FUNCTION_BLOCK basicPreparadorVibropac (* Preparador de polimero Vibropac VIB-3000 - logica (Modbus TCP Inovaisa) *)
  (* Standard: 61499-2 *)
  (* Version 1.0, 19/10/2026, Hidryco, Hidryco, 1.0: liga/desliga ciclo remoto (4001, reenvio a cada 5 s), reset 4002 por 3 s, leitura 4005..4019, modo automatico/manual, cfgHabilitada *)
  PACKAGE Hidryco.HidrycoLib;
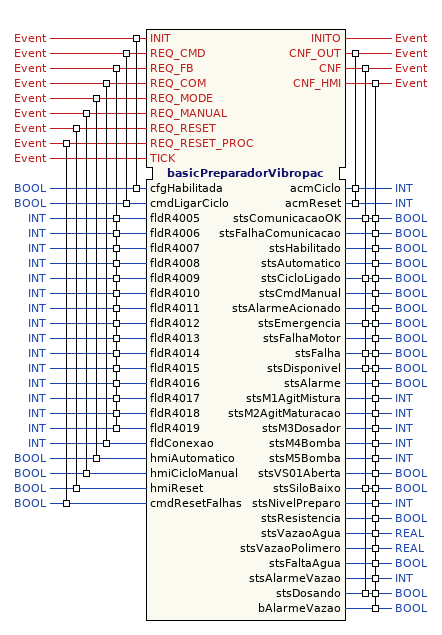
  EVENT_INPUT
    INIT WITH cfgHabilitada; (* Inicializacao (configuracao da instancia) *)
    REQ_CMD WITH cmdLigarCiclo; (* Processo: liga/desliga o ciclo (automatico) *)
    REQ_FB WITH fldR4005, fldR4006, fldR4007, fldR4008, fldR4009, fldR4010, fldR4011, fldR4012, fldR4013, fldR4014, fldR4015, fldR4016, fldR4017, fldR4018, fldR4019; (* Leitura Modbus 4005..4019 *)
    REQ_COM WITH fldConexao; (* Status da conexao Modbus (connStatusInt) *)
    REQ_MODE WITH hmiAutomatico; (* IHM: modo *)
    REQ_MANUAL WITH hmiCicloManual; (* IHM: liga/desliga o ciclo em manual *)
    REQ_RESET WITH hmiReset; (* IHM: reset *)
    REQ_RESET_PROC WITH cmdResetFalhas; (* Processo: reset *)
    TICK; (* Base de tempo de 1 s *)
  END_EVENT
  EVENT_OUTPUT
    INITO; (* Inicializacao concluida *)
    CNF_OUT WITH acmCiclo, acmReset; (* Escrita Modbus 4001 (ciclo) e 4002 (reset) *)
    CNF WITH stsComunicacaoOK, stsDisponivel, stsCicloLigado, stsFalha, stsEmergencia, stsDosando, stsSiloBaixo; (* Status para o processo (na mudanca e a cada 1 s) *)
    CNF_HMI WITH stsComunicacaoOK, stsFalhaComunicacao, stsHabilitado, stsAutomatico, stsCicloLigado, stsCmdManual, stsAlarmeAcionado, stsEmergencia, stsFalhaMotor, stsFalha, stsDisponivel, stsAlarme, stsM1AgitMistura, stsM2AgitMaturacao, stsM3Dosador, stsM4Bomba, stsM5Bomba, stsVS01Aberta, stsSiloBaixo, stsNivelPreparo, stsResistencia, stsVazaoAgua, stsVazaoPolimero, stsFaltaAgua, stsAlarmeVazao, stsDosando, bAlarmeVazao; (* Status para a IHM e alarmes *)
  END_EVENT
  VAR_INPUT
    cfgHabilitada : BOOL := TRUE; (* FALSE = instancia desabilitada (equipamento futuro): sem alarme e nunca disponivel *)
    cmdLigarCiclo : BOOL; (* Processo: TRUE = ciclo remoto ligado *)
    fldR4005 : INT; (* Registro 4005: alarme acionado (0/1) *)
    fldR4006 : INT; (* Registro 4006: emergencia (0/1) *)
    fldR4007 : INT; (* Registro 4007: status M1 agitador do tanque de mistura (0 parado, 1 funcionando, 2 falha) *)
    fldR4008 : INT; (* Registro 4008: status M2 agitador do tanque de maturacao (0 parado, 1 funcionando, 2 falha) *)
    fldR4009 : INT; (* Registro 4009: status M3 dosador volumetrico (0 parado, 1 funcionando, 2 falha) *)
    fldR4010 : INT; (* Registro 4010: status M4 bomba dosadora M4 (0 parado, 1 funcionando, 2 falha) *)
    fldR4011 : INT; (* Registro 4011: status M5 bomba dosadora M5 (0 parado, 1 funcionando, 2 falha) *)
    fldR4012 : INT; (* Registro 4012: ver tabela Modbus *)
    fldR4013 : INT; (* Registro 4013: ver tabela Modbus *)
    fldR4014 : INT; (* Registro 4014: ver tabela Modbus *)
    fldR4015 : INT; (* Registro 4015: ver tabela Modbus *)
    fldR4016 : INT; (* Registro 4016: ver tabela Modbus *)
    fldR4017 : INT; (* Registro 4017: ver tabela Modbus *)
    fldR4018 : INT; (* Registro 4018: ver tabela Modbus *)
    fldR4019 : INT; (* Registro 4019: ver tabela Modbus *)
    fldConexao : INT; (* connStatusInt (1 = online) *)
    hmiAutomatico : BOOL; (* IHM: TRUE = automatico *)
    hmiCicloManual : BOOL; (* IHM: TRUE = liga o ciclo (manual) *)
    hmiReset : BOOL; (* IHM: reset *)
    cmdResetFalhas : BOOL; (* Processo: reset (vale com TRUE) *)
  END_VAR
  VAR_OUTPUT
    acmCiclo : INT; (* Registro 4001: 1 liga ciclo remoto, 0 desliga *)
    acmReset : INT; (* Registro 4002: 1 reseta falhas (pulso de 3 s) *)
    stsComunicacaoOK : BOOL; (* Comunicacao Modbus com o CLP do skid OK *)
    stsFalhaComunicacao : BOOL; (* Falha de comunicacao com o CLP do skid *)
    stsHabilitado : BOOL; (* Instancia habilitada (FALSE = equipamento futuro) *)
    stsAutomatico : BOOL; (* Ciclo comandado pelo processo (automatico) *)
    stsCicloLigado : BOOL; (* Comando de ciclo remoto ligado (4001 = 1) *)
    stsCmdManual : BOOL; (* Comando manual de ciclo (modo manual) *)
    stsAlarmeAcionado : BOOL; (* Alarme acionado no skid (4005) *)
    stsEmergencia : BOOL; (* Botao de emergencia do skid acionado (4006) *)
    stsFalhaMotor : BOOL; (* Algum motor do skid em falha *)
    stsFalha : BOOL; (* Skid em falha (alarme, emergencia ou motor) *)
    stsDisponivel : BOOL; (* Pode ser ligado pelo automatico agora *)
    stsAlarme : BOOL; (* Algum alarme do skid *)
    stsM1AgitMistura : INT; (* Status M1 agitador do tanque de mistura (4007): 0 parado, 1 funcionando, 2 falha *)
    stsM2AgitMaturacao : INT; (* Status M2 agitador do tanque de maturacao (4008): 0 parado, 1 funcionando, 2 falha *)
    stsM3Dosador : INT; (* Status M3 dosador volumetrico (4009): 0 parado, 1 funcionando, 2 falha *)
    stsM4Bomba : INT; (* Status M4 bomba dosadora M4 (4010): 0 parado, 1 funcionando, 2 falha *)
    stsM5Bomba : INT; (* Status M5 bomba dosadora M5 (4011): 0 parado, 1 funcionando, 2 falha *)
    stsVS01Aberta : BOOL; (* Solenoide de agua VS-01 aberta (4012) *)
    stsSiloBaixo : BOOL; (* Silo de polimero em po com nivel baixo LSL-01 (4013 = 0) *)
    stsNivelPreparo : INT; (* Nivel LS1: 0 muito baixo, 1 baixo, 2 alto, 3 muito alto (4014) *)
    stsResistencia : BOOL; (* Resistencia de aquecimento RA-01 ligada (4015) *)
    stsVazaoAgua : REAL; (* Vazao de agua FIT-01 (%) (4016, 0-1000) *)
    stsVazaoPolimero : REAL; (* Vazao de polimero preparado FIT-02 (%) (4017, 0-1000) *)
    stsFaltaAgua : BOOL; (* Alarme de falta d agua (4018) *)
    stsAlarmeVazao : INT; (* Alarme de vazao de polimero: 0 sem, 1 baixa, 2 alta (4019) *)
    stsDosando : BOOL; (* Bomba dosadora M4 ou M5 funcionando *)
    bAlarmeVazao : BOOL; (* Alarme de vazao de polimero (baixa ou alta) *)
  END_VAR
  VAR
    initDone : BOOL;
    comRecebido : BOOL;
    fbRecebido : BOOL;
    bAuto : BOOL := TRUE; (* Modo automatico (partida em automatico) *)
    bFalhaMotor : BOOL;
    tReset : INT; (* Segundos restantes do pulso de reset *)
    tEnvio : INT;
    oldCiclo : INT := -1;
    oldReset : INT := -1;
    primeiro : BOOL := TRUE;
    sig : INT;
    oldSig : INT := -1;
  END_VAR
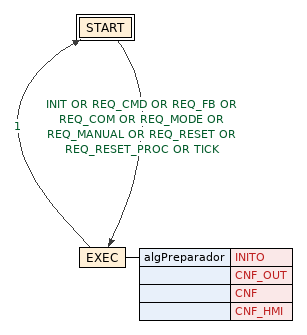
  EC_STATES
    START; (* Estado inicial *)
    EXEC : algPreparador -> INITO, -> CNF_OUT, -> CNF, -> CNF_HMI; (* Executa a logica; o algoritmo decide quais eventos saem *)
  END_STATES
  EC_TRANSITIONS
    START TO EXEC := INIT OR REQ_CMD OR REQ_FB OR REQ_COM OR REQ_MODE OR REQ_MANUAL OR REQ_RESET OR REQ_RESET_PROC OR TICK;
    EXEC TO START := 1;
  END_TRANSITIONS
  ALGORITHM algPreparador IN ST: (* Logica completa (um unico algoritmo) *)
(* =====================================================================
   basicPreparadorVibropac v1.0 - logica do CAT Preparador_Vibropac (HidrycoLib)
   Preparador de polimero Vibropac VIB-3000 - CLP do skid (M241) servidor Modbus TCP, tabela
   Inovaisa: 4001 liga/desliga ciclo remoto, 4002 reset, status a partir
   de 4005. O skid tem a propria logica (sequencia, intertravamentos e
   limpeza); o CLP da planta so liga/desliga o ciclo e le os estados.
   Regras:
   - automatico: ciclo = cmdLigarCiclo do processo; manual: comando da IHM;
   - o comando 4001 e reenviado a cada 5 s (o skid guarda o ultimo valor);
   - reset (IHM ou processo): 4002 = 1 por 3 s e reconhece os alarmes;
   - sem comunicacao: estados zerados, alarme de comunicacao (aviso);
   - cfgHabilitada = FALSE: equipamento futuro, sem alarme, ciclo desligado.
   ===================================================================== *)

INITO   := FALSE;
CNF_OUT := FALSE;
CNF     := FALSE;
CNF_HMI := FALSE;

IF REQ_COM THEN
    comRecebido := TRUE;
END_IF;
IF REQ_FB THEN
    fbRecebido := TRUE;
END_IF;
IF INIT THEN
    initDone := TRUE;
    INITO := TRUE;
END_IF;
IF NOT initDone THEN
    RETURN;
END_IF;

(* ---- 1. Comunicacao e decodificacao ---- *)
stsHabilitado := cfgHabilitada;
stsComunicacaoOK := cfgHabilitada AND comRecebido AND fbRecebido AND (fldConexao = 1);
stsFalhaComunicacao := cfgHabilitada AND NOT stsComunicacaoOK;
IF stsComunicacaoOK THEN
    stsAlarmeAcionado := fldR4005 <> 0;
    stsEmergencia := fldR4006 <> 0;
    stsM1AgitMistura := fldR4007;
    stsM2AgitMaturacao := fldR4008;
    stsM3Dosador := fldR4009;
    stsM4Bomba := fldR4010;
    stsM5Bomba := fldR4011;

    stsVS01Aberta := fldR4012 = 1;
    stsSiloBaixo := fldR4013 = 0;
    stsNivelPreparo := fldR4014;
    stsResistencia := fldR4015 = 1;
    stsVazaoAgua := LIMIT(0.0, INT_TO_REAL(fldR4016) / 10.0, 100.0);
    stsVazaoPolimero := LIMIT(0.0, INT_TO_REAL(fldR4017) / 10.0, 100.0);
    stsFaltaAgua := fldR4018 <> 0;
    stsAlarmeVazao := fldR4019;
    stsDosando := (fldR4010 = 1) OR (fldR4011 = 1);
    bFalhaMotor := (fldR4007 = 2) OR (fldR4008 = 2) OR (fldR4009 = 2) OR (fldR4010 = 2) OR (fldR4011 = 2);
ELSE
    stsAlarmeAcionado := FALSE;
    stsEmergencia := FALSE;
    stsM1AgitMistura := 0;
    stsM2AgitMaturacao := 0;
    stsM3Dosador := 0;
    stsM4Bomba := 0;
    stsM5Bomba := 0;
    stsVS01Aberta := FALSE; stsSiloBaixo := FALSE; stsResistencia := FALSE; stsFaltaAgua := FALSE; stsAlarmeVazao := 0; stsDosando := FALSE; bFalhaMotor := FALSE;
END_IF;
stsFalhaMotor := bFalhaMotor;
stsFalha := stsAlarmeAcionado OR stsEmergencia OR bFalhaMotor;
bAlarmeVazao := stsComunicacaoOK AND (stsAlarmeVazao <> 0);

(* ---- 2. Modo, comando e reset ---- *)
IF REQ_MODE THEN
    bAuto := hmiAutomatico;
END_IF;
IF REQ_MANUAL THEN
    stsCmdManual := hmiCicloManual;
END_IF;
IF bAuto THEN
    stsCmdManual := FALSE;                 (* volta ao automatico sem comando manual pendente *)
END_IF;
stsAutomatico := bAuto;
IF NOT cfgHabilitada THEN
    stsCicloLigado := FALSE;
ELSIF bAuto THEN
    stsCicloLigado := cmdLigarCiclo;
ELSE
    stsCicloLigado := stsCmdManual;
END_IF;
IF (REQ_RESET AND hmiReset) OR (REQ_RESET_PROC AND cmdResetFalhas) THEN
    tReset := 3;
END_IF;
IF TICK AND (tReset > 0) THEN
    tReset := tReset - 1;
END_IF;
IF stsCicloLigado THEN
    acmCiclo := 1;
ELSE
    acmCiclo := 0;
END_IF;
IF tReset > 0 THEN
    acmReset := 1;
ELSE
    acmReset := 0;
END_IF;
IF TICK THEN
    tEnvio := tEnvio + 1;
END_IF;
IF cfgHabilitada AND (primeiro OR (acmCiclo <> oldCiclo) OR (acmReset <> oldReset) OR (tEnvio >= 5)) THEN
    CNF_OUT := TRUE;
    tEnvio := 0;
    oldCiclo := acmCiclo;
    oldReset := acmReset;
END_IF;

(* ---- 3. Disponibilidade e alarme ---- *)
stsDisponivel := stsComunicacaoOK AND bAuto AND NOT stsFalha;
stsAlarme := stsFalhaComunicacao OR stsFalha OR stsSiloBaixo OR stsFaltaAgua OR bAlarmeVazao;

(* ---- 4. Eventos ---- *)
sig := 0;
IF stsComunicacaoOK THEN sig := sig + 1; END_IF;
IF stsDisponivel THEN sig := sig + 2; END_IF;
IF stsCicloLigado THEN sig := sig + 4; END_IF;
IF stsFalha THEN sig := sig + 8; END_IF;
IF stsEmergencia THEN sig := sig + 16; END_IF;
IF stsAlarme THEN sig := sig + 32; END_IF;
IF stsDosando THEN sig := sig + 64; END_IF;
IF bAuto THEN sig := sig + 128; END_IF;
IF primeiro OR TICK OR REQ_RESET OR REQ_MODE OR REQ_MANUAL OR (sig <> oldSig) THEN
    CNF_HMI := TRUE;
END_IF;
IF primeiro OR TICK OR (sig <> oldSig) THEN
    CNF := TRUE;
END_IF;
oldSig := sig;
primeiro := FALSE;
  END_ALGORITHM
END_FUNCTION_BLOCK
